Fanuc KAREL source: kb00062.KL

-- PROVISIONAL review KL for V1013-1; original PC SHA256 3bc91cef8d3e1762650b66ad23b305a6800d59fa97f9565f5383e5ef980a7e1d
-- Incomplete behavior may be omitted. Consult companion uncertainty JSON. Do not deploy.
PROGRAM KB00062
%NOLOCKGROUP
BEGIN
  -- UNRESOLVED_PC offsets 5-12; opcodes 9D,23
  -- UNRESOLVED_PC offsets 17-27; opcodes 9D,22,9D,33,35
  -- UNRESOLVED_PC offsets 32-39; opcodes 9D,23
  -- UNRESOLVED_PC offsets 44-72; opcodes 27,22,22,22,22,31
  -- UNRESOLVED_PC offsets 77-81; opcodes 7F
END KB00062
